Fanuc KAREL source: kd00062.KL

-- PROVISIONAL review KL for V770-1; original PC SHA256 1ea3edd5ad3a72d4cfed45b57d287c31948343dd7d982ca4fe39d95736793772
-- Incomplete behavior may be omitted. Consult companion uncertainty JSON. Do not deploy.
PROGRAM KD00062
%NOLOCKGROUP
VAR
  I : INTEGER
  J : INTEGER
  B : BOOLEAN
  R : REAL
  S : STRING[80]
BEGIN
  -- UNRESOLVED_PC offsets 5-18; opcodes 9D,81,18,9D,1B,9D,12,9D,13,04
  -- UNRESOLVED_PC offsets 23-27; opcodes 7F
END KD00062
